// TIA Portal V19 export
TYPE "EM04_Output"
   STRUCT
      Status : "EM_Output";
   END_STRUCT;
END_TYPE
